Fanuc KAREL source: KA00113.KL

PROGRAM KA00113
%NOLOCKGROUP
VAR
  SRC: CONFIG
  DST: POSITION
BEGIN
  SRC.CFG_FLIP = TRUE
  DST = SRC
END KA00113
